(*
SPDX-FileCopyrightText: © 2026 Oleksandr Tiutyk <trofimich@gmail.com>
SPDX-License-Identifier: MIT
License: https://opensource.org/license/mit
*)

(*!
<summary>Condition that inverts the evaluation result of an inner workflow condition.</summary>
<description>
Evaluates the inner condition via Evaluate and returns the logical negation of its result. Requires a
non-null, configured inner condition to be considered Configured.
</description>
*)

{attribute 'no_explicit_call' := 'do not call this function block directly'}
{attribute 'enable_dynamic_creation'}
FUNCTION_BLOCK NotCondition EXTENDS Condition IMPLEMENTS INotCondition, TOF_Core.IConfigurationSerializable
VAR_STAT
	{attribute 'hide'}
	_ClassName : STRING := __POUNAME();
END_VAR
VAR
	{attribute 'OPC.UA.DA' := '0'}
	_Condition : ICondition;
END_VAR

(*!
<summary>Borrows the initialized class name used in diagnostics.</summary>
<description>
Returns initialized metadata storage without allocation. Callers must not modify the returned string.
Derived function blocks must use distinct initialized static storage when overriding this metadata.
</description>
*)
{attribute 'monitoring' := 'call'}
PROPERTY ClassName : REFERENCE TO STRING
GET
ClassName REF= _ClassName;
END_GET
END_PROPERTY

(*!
<summary>Gets the inner condition whose evaluation result is inverted.</summary>
*)
{attribute 'monitoring' := 'call'}
PROPERTY Condition : ICondition
GET
Condition := _Condition;
END_GET
END_PROPERTY

(*!
<summary>Reports whether the inner condition has been configured and is ready for evaluation.</summary>
*)
{attribute 'monitoring' := 'call'}
PROPERTY Configured : BOOL
GET
Configured := _Condition <> 0 AND_THEN _Condition.Configured;
END_GET
END_PROPERTY

(*!
<summary>Configures the inner condition to be inverted.</summary>
<description>
Validates that the condition is not null, not this condition itself or an ancestor, and not already attached
to another parent.
The parent chain and owning workflow must be PASSIVE_READY; fixed workflow association is checked before
mutation. Reusing the same dependency is permitted. Replaced dependencies retain their existing parent links
and must not be attached elsewhere. Parent callbacks are not transactional. Dependencies remain borrowed.
</description>
<param name="condition">Inner condition to invert.</param>
*)
METHOD Configure
VAR_INPUT
	condition : ICondition;
END_VAR
ValidateConditionAttachment(condition := condition, argumentName := 'condition');

_Condition := condition;
condition.ParentCondition := THIS^;
END_METHOD

(*!
<summary>Borrows the compiler-initialized library namespace.</summary>
<description>
Borrows storage from the live internal namespace provider. Reacquire references after application
reinitialization or relocation. Treat the reference as read-only; no ownership or synchronization is provided.
</description>
*)
{attribute 'monitoring' := 'call'}
PROPERTY NamespaceName : REFERENCE TO STRING
GET
NamespaceName REF= CurrentNamespace.Name;
END_GET
END_PROPERTY

(*!
<summary>Evaluates the inner condition and returns its logical negation.</summary>
<param name="activity">Activity context for variable lookup.</param>
*)
METHOD PROTECTED OnEvaluate : BOOL
VAR_INPUT
	activity : IActivity;
END_VAR
VAR
	formattedExceptionMessage : TOF_Core.ERROR_MESSAGE;
END_VAR
IF NOT Configured THEN
	formattedExceptionMessage := TOF_Core.WideStrings.Concat255("Condition '", Name, "' is not configured");

	WorkflowExceptions.ThrowWorkflowConfiguration(
		sourceNamespaceName := NamespaceName,
		sourceClassName := ClassName,
		sourcePOUName := __POUNAME(),
		sourcePosition := __POSITION(),
		message := formattedExceptionMessage
	);
END_IF

OnEvaluate := NOT _Condition.Evaluate(activity := activity);
END_METHOD

(*!
<summary>Reports the size of this concrete function block instance in bytes.</summary>
<description>
Reports the instance layout rather than dynamic allocations owned by its fields. A derived function block
with a different layout must override this property; the value does not grant disposal rights.
</description>
*)
{attribute 'monitoring' := 'call'}
PROPERTY SelfSize : ULINT
GET
SelfSize := XSIZEOF(THIS^);
END_GET
END_PROPERTY

(*!
<summary>
Verifies that an inner condition can be attached to this negation wrapper without cycles or conflicts.
</summary>
<param name="condition">Condition candidate to validate.</param>
<param name="argumentName">Parameter name for diagnostic reporting.</param>
*)
METHOD PROTECTED ValidateConditionAttachment
VAR_INPUT
	condition : ICondition;
	argumentName : STRING(255);
END_VAR
IF condition = 0 THEN
	TOF_Core.Exceptions.ThrowArgumentNotSpecified(
		sourceNamespaceName := NamespaceName,
		sourceClassName := ClassName,
		sourcePOUName := __POUNAME(),
		sourcePosition := __POSITION(),
		argumentName := argumentName
	);
END_IF

Workflows.ValidateElementAttachment(parent := THIS^, child := condition);
END_METHOD

(*!
<summary>Writes the configuration fields for this object.</summary>
<description>Borrows the writer for this call. A failure invalidates the current output document.</description>
*)
METHOD Serialize
VAR_INPUT
	writer : TOF_Core.IConfigurationWriter;
END_VAR
Workflows.WriteConfigurationHeader(writer := writer, source := THIS^, displayName := Name, scope := THIS^);
Workflows.WriteConfigurationObject(writer := writer, name := 'condition', source := _Condition);
END_METHOD

(*!
<summary>Restores this fresh instance from its configuration object.</summary>
<description>
The reader, document node and deserialization context are borrowed for this call.
On failure discard the partial instance.
</description>
<param name="reader">Active configuration reader.</param>
<param name="node">Object node to read fields from.</param>
<param name="context">Active configuration deserialization context providing workflow reconstruction services.</param>
*)
METHOD Deserialize
VAR_INPUT
	reader : TOF_Core.IConfigurationReader;
	node : TOF_Core.CONFIGURATION_NODE;
	context : TOF_Core.IConfigurationDeserializationContext;
END_VAR
VAR
	loader : IWorkflowLoader;
END_VAR
loader := WorkflowConfigurationSerializer.ResolveWorkflowLoader(context := context);
Workflows.ReadConfigurationHeader(reader := reader, node := node, target := THIS^, scope := THIS^);

Configure(
	condition := Workflows.ReadCondition(
		loader := loader,
		node := reader.GetField(node := node, name := 'condition')
	)
);
END_METHOD

END_FUNCTION_BLOCK

(* stored: Version 1.1.0.1
   POU NotCondition: Id {07037407-734f-48fc-9bea-f1f4eb24144b}, SpecialFunc None
   Folder Overriden methods: Id {3a817429-0fa1-41b2-bf58-9a3b2167edfa}
   Folder Service methods: Id {b93590a6-dd9b-4289-bf40-a61da5548aea}
   Property ClassName: Id {bca735fa-76c8-4113-8046-d96caa463f1b}
   Get Get: Id {9ad56043-d757-444d-b758-425c6ce04d39}
   Property Condition: Id {32b77fcc-93ca-49a3-8432-613313d7a66d}
   Get Get: Id {d1f9b7a5-8a62-45ab-ad96-3f31da99c90a}
   Property Configured: Id {aacb589b-8c73-4aad-bf10-28beb66feaf1}
   Get Get: Id {2464377e-9bae-4b3f-b0f3-10e6b95ad25b}
   Method Configure: Id {abc1db78-0e72-457d-9142-b2d5a0d8938b}
   Property NamespaceName: Id {42ff9a00-beff-49d9-9666-03a047f67985}
   Get Get: Id {c12881cc-90f9-4ba4-a93d-ce9b87971edc}
   Method OnEvaluate: Id {2980fd52-bd90-48be-a8d9-65fd93889672}
   Property SelfSize: Id {52232918-81b2-434b-820c-49bd1bbcb29a}
   Get Get: Id {5565922b-1d3d-4db0-9941-176d41d9b15c}
   Method ValidateConditionAttachment: Id {5eedc3dc-858b-4e55-9016-c2022c97226c}
   Method Serialize: Id {81195d08-019b-498e-98af-cb9a3ac42f5c}
   Method Deserialize: Id {7aceabb4-b2a4-4505-b685-8becc40f6a1d} *)
